Fanuc KAREL source: compact_preamble.KL

PROGRAM KA00092
%NOLOCKGROUP
VAR
SRC : JOINTPOS9
DST : JOINTPOS9
BEGIN
DST=SRC
END KA00092
